SUBAPPLICATION Uebung_156b (* Übung zu FsGet/FsPut: Datei vom File Server holen und als Kopie zurückschreiben *)
  (* Standard: 61499-2; Description: Copyright (c) 2026 Meisterschulen am Ostbahnhof This program and the accompanying materials are made available under the terms of the Eclipse Public License 2.0 which is available at https://www.eclipse.org/legal/epl-2.0/ SPDX-License-Identifier: EPL-2.0 *)
  (* Version 1.0, 2026-11-25, Franz Höpfinger, Meisterschulen am Ostbahnhof, initial API and implementation and/or initial documentation *)
  PACKAGE Uebungen;
  IMPORT Uebungen::const::Uebung_150_159::FileServer::FS_ADD;
  IMPORT Uebungen::const::Uebung_150_159::FileServer::FS_DATEI;
  IMPORT Uebungen::const::Uebung_150_159::FileServer::FS_DATEI_2;
  IMPORT Uebungen::const::Uebung_150_159::FileServer::FS_FLT;
  IMPORT Uebungen::const::Uebung_150_159::FileServer::FS_LOKAL;
  IMPORT isobus::pgn::ISOUSERHOME_e::network;
  IMPORT isobus::pgn::ISO_CAN_NODE::NODE1;
  IMPORT logiBUS::io::DI::logiBUS_DI::Input_I1;
  IMPORT logiBUS::io::DI::logiBUS_DI_Events::BUTTON_SINGLE_CLICK;
  IMPORT logiBUS::io::DQ::logiBUS_DO::Output_Q1;
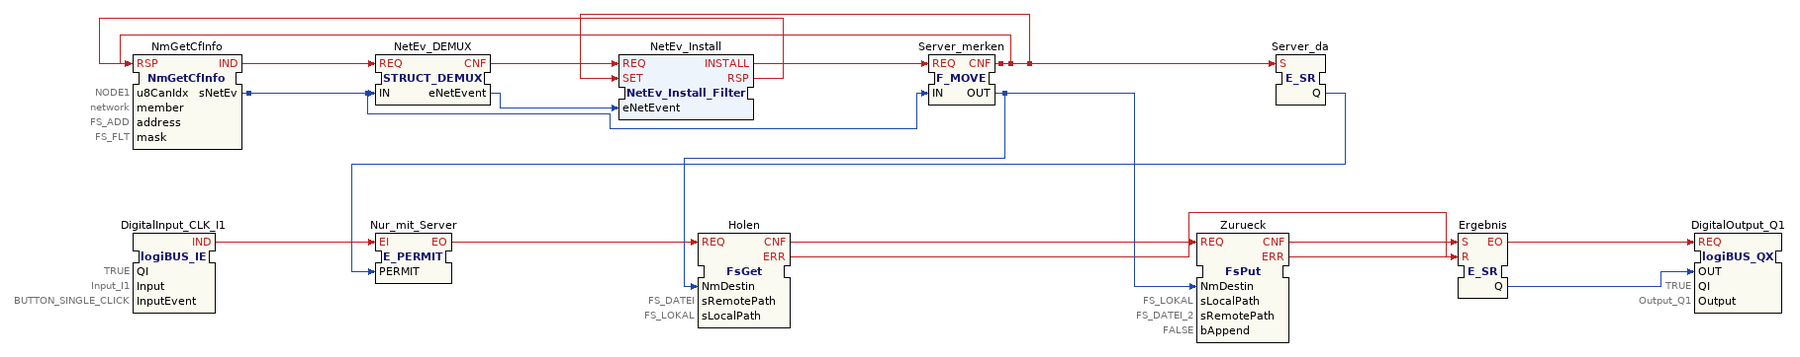
  (* File Server: Datei holen und als Kopie zurückschreiben (FsGet, FsPut) NmGetCfInfo (network, Filter FS_ADD/FS_FLT = NAME-Funktion 61) meldet den File Server, z. B. CCI 1200 mit USB-Stick. I1 Klick (nur mit Server): FS_DATEI nach FS_LOKAL (/data/fs/) holen, dann als FS_DATEI_2 zurückschreiben. Q1 an = fertig, Q1 aus = Fehler. Watch: u32Bytes (PROG beim Holen), bei ERR s16Status und u16FsError. FS_DATEI muss es geben, z. B. aus Übung 156. Voraussetzungen: Firmware ab LOGIBUS f6afe1e4 (File Server Client), isobus_fs-ELF, PART_13_FSC = 1 in /data/functionalities.ini. Lokale Pfade nur unter /data/fs/ (bei einem logiBUS als Server: /data/). *)
  FBS
    NmGetCfInfo : isobus::pgn::NmGetCfInfo(u8CanIdx := NODE1, member := network, address := FS_ADD, mask := FS_FLT); (* meldet den File Server (Funktion 61) *)
    NetEv_DEMUX : eclipse4diac::convert::STRUCT_DEMUX; {SET_ATTRIBUTE(StructuredType, isobus::pgn::ISONETEVENT_T)}
    Server_merken : iec61131::selection::F_MOVE; (* eigener CF und File-Server-CF (NmDestin) *)
    Server_da : iec61499::events::E_SR;
    DigitalInput_CLK_I1 : logiBUS::io::DI::logiBUS_IE(QI := TRUE, Input := Input_I1, InputEvent := BUTTON_SINGLE_CLICK);
    Nur_mit_Server : iec61499::events::E_PERMIT;
    Holen : isobus::fs::FsGet(sRemotePath := FS_DATEI, sLocalPath := FS_LOKAL); (* FS_DATEI nach FS_LOKAL (/data/fs/...) *)
    Zurueck : isobus::fs::FsPut(sLocalPath := FS_LOKAL, sRemotePath := FS_DATEI_2, bAppend := FALSE); (* FS_LOKAL als FS_DATEI_2 zurück *)
    Ergebnis : iec61499::events::E_SR; (* Q1 an = beide Kopien fertig *)
    DigitalOutput_Q1 : logiBUS::io::DQ::logiBUS_QX(QI := TRUE, Output := Output_Q1);
  END_FBS
  SUBAPPS
    NetEv_Install : MyLib::sys::NetEv_Install_Filter;
  END_SUBAPPS
  EVENT_CONNECTIONS
    NmGetCfInfo.IND TO NetEv_DEMUX.REQ;
    NetEv_DEMUX.CNF TO NetEv_Install.REQ;
    NetEv_Install.INSTALL TO Server_merken.REQ;
    NetEv_Install.RSP TO NmGetCfInfo.RSP;
    Server_merken.CNF TO NetEv_Install.SET;
    Server_merken.CNF TO Server_da.S;
    Server_merken.CNF TO NmGetCfInfo.RSP;
    DigitalInput_CLK_I1.IND TO Nur_mit_Server.EI;
    Nur_mit_Server.EO TO Holen.REQ;
    Holen.CNF TO Zurueck.REQ;
    Zurueck.CNF TO Ergebnis.S;
    Holen.ERR TO Ergebnis.R;
    Zurueck.ERR TO Ergebnis.R;
    Ergebnis.EO TO DigitalOutput_Q1.REQ;
  END_CONNECTIONS
  DATA_CONNECTIONS
    NmGetCfInfo.sNetEv TO NetEv_DEMUX.IN;
    NetEv_DEMUX.eNetEvent TO NetEv_Install.eNetEvent;
    NmGetCfInfo.sNetEv TO Server_merken.IN;
    Server_merken.OUT TO Holen.NmDestin;
    Server_merken.OUT TO Zurueck.NmDestin;
    Server_da.Q TO Nur_mit_Server.PERMIT;
    Ergebnis.Q TO DigitalOutput_Q1.OUT;
  END_CONNECTIONS
END_SUBAPPLICATION
